(* IEC 61131-3 sources: STAR-PLC-Agent/results/raw/six_task_fullflow_20261114/PUB016/generation/sim_00, 1 file *)

(* ---- test_program.st ---- *)
PROGRAM PLC_PRG
VAR
 BenchStep : UDINT := 0;
 BenchCalls : UDINT := 0;
 BenchDone : BOOL := FALSE;
 BenchUut0 : FB_Task;
 BenchUut1 : FB_Task;
 TraceIn_processLength : ARRAY[0..12] OF USINT;
 TraceIn_sensor1 : ARRAY[0..12] OF BOOL;
 TraceIn_sensor2 : ARRAY[0..12] OF BOOL;
 TraceIn_sensor3 : ARRAY[0..12] OF BOOL;
 TraceIn_sensor4 : ARRAY[0..12] OF BOOL;
 TraceIn_sensor5 : ARRAY[0..12] OF BOOL;
 TraceIn_station1Start : ARRAY[0..12] OF BOOL;
 TraceIn_station2Complete : ARRAY[0..12] OF BOOL;
 TraceIn_station3Complete : ARRAY[0..12] OF BOOL;
 TraceIn_station4Complete : ARRAY[0..12] OF BOOL;
 TraceIn_processSequence_1 : ARRAY[0..12] OF USINT;
 TraceIn_processSequence_2 : ARRAY[0..12] OF USINT;
 TraceIn_processSequence_3 : ARRAY[0..12] OF USINT;
 TraceIn_processSequence_4 : ARRAY[0..12] OF USINT;
 TraceIn_processSequence_5 : ARRAY[0..12] OF USINT;
 TraceIn_processSequence_6 : ARRAY[0..12] OF USINT;
 TraceIn_processSequence_7 : ARRAY[0..12] OF USINT;
 TraceIn_processSequence_8 : ARRAY[0..12] OF USINT;
 TraceOut_conveyorLeft : ARRAY[0..12] OF BOOL;
 TraceOut_conveyorRight : ARRAY[0..12] OF BOOL;
END_VAR

IF NOT BenchDone THEN
 CASE BenchStep OF
 0:
   BenchUut0.processLength := USINT#2;
   BenchUut0.sensor1 := TRUE;
   BenchUut0.sensor2 := FALSE;
   BenchUut0.sensor3 := FALSE;
   BenchUut0.sensor4 := FALSE;
   BenchUut0.sensor5 := FALSE;
   BenchUut0.station1Start := FALSE;
   BenchUut0.station2Complete := FALSE;
   BenchUut0.station3Complete := FALSE;
   BenchUut0.station4Complete := FALSE;
   BenchUut0.processSequence[1] := USINT#2;
   BenchUut0.processSequence[2] := USINT#5;
   BenchUut0.processSequence[3] := USINT#0;
   BenchUut0.processSequence[4] := USINT#0;
   BenchUut0.processSequence[5] := USINT#0;
   BenchUut0.processSequence[6] := USINT#0;
   BenchUut0.processSequence[7] := USINT#0;
   BenchUut0.processSequence[8] := USINT#0;
   TraceIn_processLength[0] := BenchUut0.processLength;
   TraceIn_sensor1[0] := BenchUut0.sensor1;
   TraceIn_sensor2[0] := BenchUut0.sensor2;
   TraceIn_sensor3[0] := BenchUut0.sensor3;
   TraceIn_sensor4[0] := BenchUut0.sensor4;
   TraceIn_sensor5[0] := BenchUut0.sensor5;
   TraceIn_station1Start[0] := BenchUut0.station1Start;
   TraceIn_station2Complete[0] := BenchUut0.station2Complete;
   TraceIn_station3Complete[0] := BenchUut0.station3Complete;
   TraceIn_station4Complete[0] := BenchUut0.station4Complete;
   TraceIn_processSequence_1[0] := BenchUut0.processSequence[1];
   TraceIn_processSequence_2[0] := BenchUut0.processSequence[2];
   TraceIn_processSequence_3[0] := BenchUut0.processSequence[3];
   TraceIn_processSequence_4[0] := BenchUut0.processSequence[4];
   TraceIn_processSequence_5[0] := BenchUut0.processSequence[5];
   TraceIn_processSequence_6[0] := BenchUut0.processSequence[6];
   TraceIn_processSequence_7[0] := BenchUut0.processSequence[7];
   TraceIn_processSequence_8[0] := BenchUut0.processSequence[8];
   BenchUut0();
   TraceOut_conveyorLeft[0] := BenchUut0.conveyorLeft;
   TraceOut_conveyorRight[0] := BenchUut0.conveyorRight;
   BenchCalls := BenchCalls + 1;
 1:
   BenchUut0.processLength := USINT#2;
   BenchUut0.sensor1 := TRUE;
   BenchUut0.sensor2 := FALSE;
   BenchUut0.sensor3 := FALSE;
   BenchUut0.sensor4 := FALSE;
   BenchUut0.sensor5 := FALSE;
   BenchUut0.station1Start := TRUE;
   BenchUut0.station2Complete := FALSE;
   BenchUut0.station3Complete := FALSE;
   BenchUut0.station4Complete := FALSE;
   BenchUut0.processSequence[1] := USINT#2;
   BenchUut0.processSequence[2] := USINT#5;
   BenchUut0.processSequence[3] := USINT#0;
   BenchUut0.processSequence[4] := USINT#0;
   BenchUut0.processSequence[5] := USINT#0;
   BenchUut0.processSequence[6] := USINT#0;
   BenchUut0.processSequence[7] := USINT#0;
   BenchUut0.processSequence[8] := USINT#0;
   TraceIn_processLength[1] := BenchUut0.processLength;
   TraceIn_sensor1[1] := BenchUut0.sensor1;
   TraceIn_sensor2[1] := BenchUut0.sensor2;
   TraceIn_sensor3[1] := BenchUut0.sensor3;
   TraceIn_sensor4[1] := BenchUut0.sensor4;
   TraceIn_sensor5[1] := BenchUut0.sensor5;
   TraceIn_station1Start[1] := BenchUut0.station1Start;
   TraceIn_station2Complete[1] := BenchUut0.station2Complete;
   TraceIn_station3Complete[1] := BenchUut0.station3Complete;
   TraceIn_station4Complete[1] := BenchUut0.station4Complete;
   TraceIn_processSequence_1[1] := BenchUut0.processSequence[1];
   TraceIn_processSequence_2[1] := BenchUut0.processSequence[2];
   TraceIn_processSequence_3[1] := BenchUut0.processSequence[3];
   TraceIn_processSequence_4[1] := BenchUut0.processSequence[4];
   TraceIn_processSequence_5[1] := BenchUut0.processSequence[5];
   TraceIn_processSequence_6[1] := BenchUut0.processSequence[6];
   TraceIn_processSequence_7[1] := BenchUut0.processSequence[7];
   TraceIn_processSequence_8[1] := BenchUut0.processSequence[8];
   BenchUut0();
   TraceOut_conveyorLeft[1] := BenchUut0.conveyorLeft;
   TraceOut_conveyorRight[1] := BenchUut0.conveyorRight;
   BenchCalls := BenchCalls + 1;
 2:
   BenchUut0.processLength := USINT#2;
   BenchUut0.sensor1 := TRUE;
   BenchUut0.sensor2 := TRUE;
   BenchUut0.sensor3 := FALSE;
   BenchUut0.sensor4 := FALSE;
   BenchUut0.sensor5 := FALSE;
   BenchUut0.station1Start := FALSE;
   BenchUut0.station2Complete := FALSE;
   BenchUut0.station3Complete := FALSE;
   BenchUut0.station4Complete := FALSE;
   BenchUut0.processSequence[1] := USINT#2;
   BenchUut0.processSequence[2] := USINT#5;
   BenchUut0.processSequence[3] := USINT#0;
   BenchUut0.processSequence[4] := USINT#0;
   BenchUut0.processSequence[5] := USINT#0;
   BenchUut0.processSequence[6] := USINT#0;
   BenchUut0.processSequence[7] := USINT#0;
   BenchUut0.processSequence[8] := USINT#0;
   TraceIn_processLength[2] := BenchUut0.processLength;
   TraceIn_sensor1[2] := BenchUut0.sensor1;
   TraceIn_sensor2[2] := BenchUut0.sensor2;
   TraceIn_sensor3[2] := BenchUut0.sensor3;
   TraceIn_sensor4[2] := BenchUut0.sensor4;
   TraceIn_sensor5[2] := BenchUut0.sensor5;
   TraceIn_station1Start[2] := BenchUut0.station1Start;
   TraceIn_station2Complete[2] := BenchUut0.station2Complete;
   TraceIn_station3Complete[2] := BenchUut0.station3Complete;
   TraceIn_station4Complete[2] := BenchUut0.station4Complete;
   TraceIn_processSequence_1[2] := BenchUut0.processSequence[1];
   TraceIn_processSequence_2[2] := BenchUut0.processSequence[2];
   TraceIn_processSequence_3[2] := BenchUut0.processSequence[3];
   TraceIn_processSequence_4[2] := BenchUut0.processSequence[4];
   TraceIn_processSequence_5[2] := BenchUut0.processSequence[5];
   TraceIn_processSequence_6[2] := BenchUut0.processSequence[6];
   TraceIn_processSequence_7[2] := BenchUut0.processSequence[7];
   TraceIn_processSequence_8[2] := BenchUut0.processSequence[8];
   BenchUut0();
   TraceOut_conveyorLeft[2] := BenchUut0.conveyorLeft;
   TraceOut_conveyorRight[2] := BenchUut0.conveyorRight;
   BenchCalls := BenchCalls + 1;
 3:
   BenchUut0.processLength := USINT#2;
   BenchUut0.sensor1 := TRUE;
   BenchUut0.sensor2 := TRUE;
   BenchUut0.sensor3 := FALSE;
   BenchUut0.sensor4 := FALSE;
   BenchUut0.sensor5 := FALSE;
   BenchUut0.station1Start := FALSE;
   BenchUut0.station2Complete := TRUE;
   BenchUut0.station3Complete := FALSE;
   BenchUut0.station4Complete := FALSE;
   BenchUut0.processSequence[1] := USINT#2;
   BenchUut0.processSequence[2] := USINT#5;
   BenchUut0.processSequence[3] := USINT#0;
   BenchUut0.processSequence[4] := USINT#0;
   BenchUut0.processSequence[5] := USINT#0;
   BenchUut0.processSequence[6] := USINT#0;
   BenchUut0.processSequence[7] := USINT#0;
   BenchUut0.processSequence[8] := USINT#0;
   TraceIn_processLength[3] := BenchUut0.processLength;
   TraceIn_sensor1[3] := BenchUut0.sensor1;
   TraceIn_sensor2[3] := BenchUut0.sensor2;
   TraceIn_sensor3[3] := BenchUut0.sensor3;
   TraceIn_sensor4[3] := BenchUut0.sensor4;
   TraceIn_sensor5[3] := BenchUut0.sensor5;
   TraceIn_station1Start[3] := BenchUut0.station1Start;
   TraceIn_station2Complete[3] := BenchUut0.station2Complete;
   TraceIn_station3Complete[3] := BenchUut0.station3Complete;
   TraceIn_station4Complete[3] := BenchUut0.station4Complete;
   TraceIn_processSequence_1[3] := BenchUut0.processSequence[1];
   TraceIn_processSequence_2[3] := BenchUut0.processSequence[2];
   TraceIn_processSequence_3[3] := BenchUut0.processSequence[3];
   TraceIn_processSequence_4[3] := BenchUut0.processSequence[4];
   TraceIn_processSequence_5[3] := BenchUut0.processSequence[5];
   TraceIn_processSequence_6[3] := BenchUut0.processSequence[6];
   TraceIn_processSequence_7[3] := BenchUut0.processSequence[7];
   TraceIn_processSequence_8[3] := BenchUut0.processSequence[8];
   BenchUut0();
   TraceOut_conveyorLeft[3] := BenchUut0.conveyorLeft;
   TraceOut_conveyorRight[3] := BenchUut0.conveyorRight;
   BenchCalls := BenchCalls + 1;
 4:
   BenchUut0.processLength := USINT#2;
   BenchUut0.sensor1 := FALSE;
   BenchUut0.sensor2 := FALSE;
   BenchUut0.sensor3 := FALSE;
   BenchUut0.sensor4 := FALSE;
   BenchUut0.sensor5 := FALSE;
   BenchUut0.station1Start := FALSE;
   BenchUut0.station2Complete := FALSE;
   BenchUut0.station3Complete := FALSE;
   BenchUut0.station4Complete := FALSE;
   BenchUut0.processSequence[1] := USINT#2;
   BenchUut0.processSequence[2] := USINT#5;
   BenchUut0.processSequence[3] := USINT#0;
   BenchUut0.processSequence[4] := USINT#0;
   BenchUut0.processSequence[5] := USINT#0;
   BenchUut0.processSequence[6] := USINT#0;
   BenchUut0.processSequence[7] := USINT#0;
   BenchUut0.processSequence[8] := USINT#0;
   TraceIn_processLength[4] := BenchUut0.processLength;
   TraceIn_sensor1[4] := BenchUut0.sensor1;
   TraceIn_sensor2[4] := BenchUut0.sensor2;
   TraceIn_sensor3[4] := BenchUut0.sensor3;
   TraceIn_sensor4[4] := BenchUut0.sensor4;
   TraceIn_sensor5[4] := BenchUut0.sensor5;
   TraceIn_station1Start[4] := BenchUut0.station1Start;
   TraceIn_station2Complete[4] := BenchUut0.station2Complete;
   TraceIn_station3Complete[4] := BenchUut0.station3Complete;
   TraceIn_station4Complete[4] := BenchUut0.station4Complete;
   TraceIn_processSequence_1[4] := BenchUut0.processSequence[1];
   TraceIn_processSequence_2[4] := BenchUut0.processSequence[2];
   TraceIn_processSequence_3[4] := BenchUut0.processSequence[3];
   TraceIn_processSequence_4[4] := BenchUut0.processSequence[4];
   TraceIn_processSequence_5[4] := BenchUut0.processSequence[5];
   TraceIn_processSequence_6[4] := BenchUut0.processSequence[6];
   TraceIn_processSequence_7[4] := BenchUut0.processSequence[7];
   TraceIn_processSequence_8[4] := BenchUut0.processSequence[8];
   BenchUut0();
   TraceOut_conveyorLeft[4] := BenchUut0.conveyorLeft;
   TraceOut_conveyorRight[4] := BenchUut0.conveyorRight;
   BenchCalls := BenchCalls + 1;
 5:
   BenchUut0.processLength := USINT#2;
   BenchUut0.sensor1 := FALSE;
   BenchUut0.sensor2 := FALSE;
   BenchUut0.sensor3 := FALSE;
   BenchUut0.sensor4 := FALSE;
   BenchUut0.sensor5 := TRUE;
   BenchUut0.station1Start := FALSE;
   BenchUut0.station2Complete := FALSE;
   BenchUut0.station3Complete := FALSE;
   BenchUut0.station4Complete := FALSE;
   BenchUut0.processSequence[1] := USINT#2;
   BenchUut0.processSequence[2] := USINT#5;
   BenchUut0.processSequence[3] := USINT#0;
   BenchUut0.processSequence[4] := USINT#0;
   BenchUut0.processSequence[5] := USINT#0;
   BenchUut0.processSequence[6] := USINT#0;
   BenchUut0.processSequence[7] := USINT#0;
   BenchUut0.processSequence[8] := USINT#0;
   TraceIn_processLength[5] := BenchUut0.processLength;
   TraceIn_sensor1[5] := BenchUut0.sensor1;
   TraceIn_sensor2[5] := BenchUut0.sensor2;
   TraceIn_sensor3[5] := BenchUut0.sensor3;
   TraceIn_sensor4[5] := BenchUut0.sensor4;
   TraceIn_sensor5[5] := BenchUut0.sensor5;
   TraceIn_station1Start[5] := BenchUut0.station1Start;
   TraceIn_station2Complete[5] := BenchUut0.station2Complete;
   TraceIn_station3Complete[5] := BenchUut0.station3Complete;
   TraceIn_station4Complete[5] := BenchUut0.station4Complete;
   TraceIn_processSequence_1[5] := BenchUut0.processSequence[1];
   TraceIn_processSequence_2[5] := BenchUut0.processSequence[2];
   TraceIn_processSequence_3[5] := BenchUut0.processSequence[3];
   TraceIn_processSequence_4[5] := BenchUut0.processSequence[4];
   TraceIn_processSequence_5[5] := BenchUut0.processSequence[5];
   TraceIn_processSequence_6[5] := BenchUut0.processSequence[6];
   TraceIn_processSequence_7[5] := BenchUut0.processSequence[7];
   TraceIn_processSequence_8[5] := BenchUut0.processSequence[8];
   BenchUut0();
   TraceOut_conveyorLeft[5] := BenchUut0.conveyorLeft;
   TraceOut_conveyorRight[5] := BenchUut0.conveyorRight;
   BenchCalls := BenchCalls + 1;
 6:
   BenchUut1.processLength := USINT#3;
   BenchUut1.sensor1 := TRUE;
   BenchUut1.sensor2 := FALSE;
   BenchUut1.sensor3 := FALSE;
   BenchUut1.sensor4 := FALSE;
   BenchUut1.sensor5 := FALSE;
   BenchUut1.station1Start := FALSE;
   BenchUut1.station2Complete := FALSE;
   BenchUut1.station3Complete := FALSE;
   BenchUut1.station4Complete := FALSE;
   BenchUut1.processSequence[1] := USINT#2;
   BenchUut1.processSequence[2] := USINT#2;
   BenchUut1.processSequence[3] := USINT#5;
   BenchUut1.processSequence[4] := USINT#0;
   BenchUut1.processSequence[5] := USINT#0;
   BenchUut1.processSequence[6] := USINT#0;
   BenchUut1.processSequence[7] := USINT#0;
   BenchUut1.processSequence[8] := USINT#0;
   TraceIn_processLength[6] := BenchUut1.processLength;
   TraceIn_sensor1[6] := BenchUut1.sensor1;
   TraceIn_sensor2[6] := BenchUut1.sensor2;
   TraceIn_sensor3[6] := BenchUut1.sensor3;
   TraceIn_sensor4[6] := BenchUut1.sensor4;
   TraceIn_sensor5[6] := BenchUut1.sensor5;
   TraceIn_station1Start[6] := BenchUut1.station1Start;
   TraceIn_station2Complete[6] := BenchUut1.station2Complete;
   TraceIn_station3Complete[6] := BenchUut1.station3Complete;
   TraceIn_station4Complete[6] := BenchUut1.station4Complete;
   TraceIn_processSequence_1[6] := BenchUut1.processSequence[1];
   TraceIn_processSequence_2[6] := BenchUut1.processSequence[2];
   TraceIn_processSequence_3[6] := BenchUut1.processSequence[3];
   TraceIn_processSequence_4[6] := BenchUut1.processSequence[4];
   TraceIn_processSequence_5[6] := BenchUut1.processSequence[5];
   TraceIn_processSequence_6[6] := BenchUut1.processSequence[6];
   TraceIn_processSequence_7[6] := BenchUut1.processSequence[7];
   TraceIn_processSequence_8[6] := BenchUut1.processSequence[8];
   BenchUut1();
   TraceOut_conveyorLeft[6] := BenchUut1.conveyorLeft;
   TraceOut_conveyorRight[6] := BenchUut1.conveyorRight;
   BenchCalls := BenchCalls + 1;
 7:
   BenchUut1.processLength := USINT#3;
   BenchUut1.sensor1 := TRUE;
   BenchUut1.sensor2 := FALSE;
   BenchUut1.sensor3 := FALSE;
   BenchUut1.sensor4 := FALSE;
   BenchUut1.sensor5 := FALSE;
   BenchUut1.station1Start := TRUE;
   BenchUut1.station2Complete := FALSE;
   BenchUut1.station3Complete := FALSE;
   BenchUut1.station4Complete := FALSE;
   BenchUut1.processSequence[1] := USINT#2;
   BenchUut1.processSequence[2] := USINT#2;
   BenchUut1.processSequence[3] := USINT#5;
   BenchUut1.processSequence[4] := USINT#0;
   BenchUut1.processSequence[5] := USINT#0;
   BenchUut1.processSequence[6] := USINT#0;
   BenchUut1.processSequence[7] := USINT#0;
   BenchUut1.processSequence[8] := USINT#0;
   TraceIn_processLength[7] := BenchUut1.processLength;
   TraceIn_sensor1[7] := BenchUut1.sensor1;
   TraceIn_sensor2[7] := BenchUut1.sensor2;
   TraceIn_sensor3[7] := BenchUut1.sensor3;
   TraceIn_sensor4[7] := BenchUut1.sensor4;
   TraceIn_sensor5[7] := BenchUut1.sensor5;
   TraceIn_station1Start[7] := BenchUut1.station1Start;
   TraceIn_station2Complete[7] := BenchUut1.station2Complete;
   TraceIn_station3Complete[7] := BenchUut1.station3Complete;
   TraceIn_station4Complete[7] := BenchUut1.station4Complete;
   TraceIn_processSequence_1[7] := BenchUut1.processSequence[1];
   TraceIn_processSequence_2[7] := BenchUut1.processSequence[2];
   TraceIn_processSequence_3[7] := BenchUut1.processSequence[3];
   TraceIn_processSequence_4[7] := BenchUut1.processSequence[4];
   TraceIn_processSequence_5[7] := BenchUut1.processSequence[5];
   TraceIn_processSequence_6[7] := BenchUut1.processSequence[6];
   TraceIn_processSequence_7[7] := BenchUut1.processSequence[7];
   TraceIn_processSequence_8[7] := BenchUut1.processSequence[8];
   BenchUut1();
   TraceOut_conveyorLeft[7] := BenchUut1.conveyorLeft;
   TraceOut_conveyorRight[7] := BenchUut1.conveyorRight;
   BenchCalls := BenchCalls + 1;
 8:
   BenchUut1.processLength := USINT#3;
   BenchUut1.sensor1 := TRUE;
   BenchUut1.sensor2 := TRUE;
   BenchUut1.sensor3 := FALSE;
   BenchUut1.sensor4 := FALSE;
   BenchUut1.sensor5 := FALSE;
   BenchUut1.station1Start := FALSE;
   BenchUut1.station2Complete := FALSE;
   BenchUut1.station3Complete := FALSE;
   BenchUut1.station4Complete := FALSE;
   BenchUut1.processSequence[1] := USINT#2;
   BenchUut1.processSequence[2] := USINT#2;
   BenchUut1.processSequence[3] := USINT#5;
   BenchUut1.processSequence[4] := USINT#0;
   BenchUut1.processSequence[5] := USINT#0;
   BenchUut1.processSequence[6] := USINT#0;
   BenchUut1.processSequence[7] := USINT#0;
   BenchUut1.processSequence[8] := USINT#0;
   TraceIn_processLength[8] := BenchUut1.processLength;
   TraceIn_sensor1[8] := BenchUut1.sensor1;
   TraceIn_sensor2[8] := BenchUut1.sensor2;
   TraceIn_sensor3[8] := BenchUut1.sensor3;
   TraceIn_sensor4[8] := BenchUut1.sensor4;
   TraceIn_sensor5[8] := BenchUut1.sensor5;
   TraceIn_station1Start[8] := BenchUut1.station1Start;
   TraceIn_station2Complete[8] := BenchUut1.station2Complete;
   TraceIn_station3Complete[8] := BenchUut1.station3Complete;
   TraceIn_station4Complete[8] := BenchUut1.station4Complete;
   TraceIn_processSequence_1[8] := BenchUut1.processSequence[1];
   TraceIn_processSequence_2[8] := BenchUut1.processSequence[2];
   TraceIn_processSequence_3[8] := BenchUut1.processSequence[3];
   TraceIn_processSequence_4[8] := BenchUut1.processSequence[4];
   TraceIn_processSequence_5[8] := BenchUut1.processSequence[5];
   TraceIn_processSequence_6[8] := BenchUut1.processSequence[6];
   TraceIn_processSequence_7[8] := BenchUut1.processSequence[7];
   TraceIn_processSequence_8[8] := BenchUut1.processSequence[8];
   BenchUut1();
   TraceOut_conveyorLeft[8] := BenchUut1.conveyorLeft;
   TraceOut_conveyorRight[8] := BenchUut1.conveyorRight;
   BenchCalls := BenchCalls + 1;
 9:
   BenchUut1.processLength := USINT#3;
   BenchUut1.sensor1 := TRUE;
   BenchUut1.sensor2 := TRUE;
   BenchUut1.sensor3 := FALSE;
   BenchUut1.sensor4 := FALSE;
   BenchUut1.sensor5 := FALSE;
   BenchUut1.station1Start := FALSE;
   BenchUut1.station2Complete := TRUE;
   BenchUut1.station3Complete := FALSE;
   BenchUut1.station4Complete := FALSE;
   BenchUut1.processSequence[1] := USINT#2;
   BenchUut1.processSequence[2] := USINT#2;
   BenchUut1.processSequence[3] := USINT#5;
   BenchUut1.processSequence[4] := USINT#0;
   BenchUut1.processSequence[5] := USINT#0;
   BenchUut1.processSequence[6] := USINT#0;
   BenchUut1.processSequence[7] := USINT#0;
   BenchUut1.processSequence[8] := USINT#0;
   TraceIn_processLength[9] := BenchUut1.processLength;
   TraceIn_sensor1[9] := BenchUut1.sensor1;
   TraceIn_sensor2[9] := BenchUut1.sensor2;
   TraceIn_sensor3[9] := BenchUut1.sensor3;
   TraceIn_sensor4[9] := BenchUut1.sensor4;
   TraceIn_sensor5[9] := BenchUut1.sensor5;
   TraceIn_station1Start[9] := BenchUut1.station1Start;
   TraceIn_station2Complete[9] := BenchUut1.station2Complete;
   TraceIn_station3Complete[9] := BenchUut1.station3Complete;
   TraceIn_station4Complete[9] := BenchUut1.station4Complete;
   TraceIn_processSequence_1[9] := BenchUut1.processSequence[1];
   TraceIn_processSequence_2[9] := BenchUut1.processSequence[2];
   TraceIn_processSequence_3[9] := BenchUut1.processSequence[3];
   TraceIn_processSequence_4[9] := BenchUut1.processSequence[4];
   TraceIn_processSequence_5[9] := BenchUut1.processSequence[5];
   TraceIn_processSequence_6[9] := BenchUut1.processSequence[6];
   TraceIn_processSequence_7[9] := BenchUut1.processSequence[7];
   TraceIn_processSequence_8[9] := BenchUut1.processSequence[8];
   BenchUut1();
   TraceOut_conveyorLeft[9] := BenchUut1.conveyorLeft;
   TraceOut_conveyorRight[9] := BenchUut1.conveyorRight;
   BenchCalls := BenchCalls + 1;
 10:
   BenchUut1.processLength := USINT#3;
   BenchUut1.sensor1 := TRUE;
   BenchUut1.sensor2 := TRUE;
   BenchUut1.sensor3 := FALSE;
   BenchUut1.sensor4 := FALSE;
   BenchUut1.sensor5 := FALSE;
   BenchUut1.station1Start := FALSE;
   BenchUut1.station2Complete := FALSE;
   BenchUut1.station3Complete := FALSE;
   BenchUut1.station4Complete := FALSE;
   BenchUut1.processSequence[1] := USINT#2;
   BenchUut1.processSequence[2] := USINT#2;
   BenchUut1.processSequence[3] := USINT#5;
   BenchUut1.processSequence[4] := USINT#0;
   BenchUut1.processSequence[5] := USINT#0;
   BenchUut1.processSequence[6] := USINT#0;
   BenchUut1.processSequence[7] := USINT#0;
   BenchUut1.processSequence[8] := USINT#0;
   TraceIn_processLength[10] := BenchUut1.processLength;
   TraceIn_sensor1[10] := BenchUut1.sensor1;
   TraceIn_sensor2[10] := BenchUut1.sensor2;
   TraceIn_sensor3[10] := BenchUut1.sensor3;
   TraceIn_sensor4[10] := BenchUut1.sensor4;
   TraceIn_sensor5[10] := BenchUut1.sensor5;
   TraceIn_station1Start[10] := BenchUut1.station1Start;
   TraceIn_station2Complete[10] := BenchUut1.station2Complete;
   TraceIn_station3Complete[10] := BenchUut1.station3Complete;
   TraceIn_station4Complete[10] := BenchUut1.station4Complete;
   TraceIn_processSequence_1[10] := BenchUut1.processSequence[1];
   TraceIn_processSequence_2[10] := BenchUut1.processSequence[2];
   TraceIn_processSequence_3[10] := BenchUut1.processSequence[3];
   TraceIn_processSequence_4[10] := BenchUut1.processSequence[4];
   TraceIn_processSequence_5[10] := BenchUut1.processSequence[5];
   TraceIn_processSequence_6[10] := BenchUut1.processSequence[6];
   TraceIn_processSequence_7[10] := BenchUut1.processSequence[7];
   TraceIn_processSequence_8[10] := BenchUut1.processSequence[8];
   BenchUut1();
   TraceOut_conveyorLeft[10] := BenchUut1.conveyorLeft;
   TraceOut_conveyorRight[10] := BenchUut1.conveyorRight;
   BenchCalls := BenchCalls + 1;
 11:
   BenchUut1.processLength := USINT#3;
   BenchUut1.sensor1 := TRUE;
   BenchUut1.sensor2 := TRUE;
   BenchUut1.sensor3 := FALSE;
   BenchUut1.sensor4 := FALSE;
   BenchUut1.sensor5 := FALSE;
   BenchUut1.station1Start := FALSE;
   BenchUut1.station2Complete := TRUE;
   BenchUut1.station3Complete := FALSE;
   BenchUut1.station4Complete := FALSE;
   BenchUut1.processSequence[1] := USINT#2;
   BenchUut1.processSequence[2] := USINT#2;
   BenchUut1.processSequence[3] := USINT#5;
   BenchUut1.processSequence[4] := USINT#0;
   BenchUut1.processSequence[5] := USINT#0;
   BenchUut1.processSequence[6] := USINT#0;
   BenchUut1.processSequence[7] := USINT#0;
   BenchUut1.processSequence[8] := USINT#0;
   TraceIn_processLength[11] := BenchUut1.processLength;
   TraceIn_sensor1[11] := BenchUut1.sensor1;
   TraceIn_sensor2[11] := BenchUut1.sensor2;
   TraceIn_sensor3[11] := BenchUut1.sensor3;
   TraceIn_sensor4[11] := BenchUut1.sensor4;
   TraceIn_sensor5[11] := BenchUut1.sensor5;
   TraceIn_station1Start[11] := BenchUut1.station1Start;
   TraceIn_station2Complete[11] := BenchUut1.station2Complete;
   TraceIn_station3Complete[11] := BenchUut1.station3Complete;
   TraceIn_station4Complete[11] := BenchUut1.station4Complete;
   TraceIn_processSequence_1[11] := BenchUut1.processSequence[1];
   TraceIn_processSequence_2[11] := BenchUut1.processSequence[2];
   TraceIn_processSequence_3[11] := BenchUut1.processSequence[3];
   TraceIn_processSequence_4[11] := BenchUut1.processSequence[4];
   TraceIn_processSequence_5[11] := BenchUut1.processSequence[5];
   TraceIn_processSequence_6[11] := BenchUut1.processSequence[6];
   TraceIn_processSequence_7[11] := BenchUut1.processSequence[7];
   TraceIn_processSequence_8[11] := BenchUut1.processSequence[8];
   BenchUut1();
   TraceOut_conveyorLeft[11] := BenchUut1.conveyorLeft;
   TraceOut_conveyorRight[11] := BenchUut1.conveyorRight;
   BenchCalls := BenchCalls + 1;
 12:
   BenchUut1.processLength := USINT#3;
   BenchUut1.sensor1 := FALSE;
   BenchUut1.sensor2 := FALSE;
   BenchUut1.sensor3 := FALSE;
   BenchUut1.sensor4 := FALSE;
   BenchUut1.sensor5 := TRUE;
   BenchUut1.station1Start := FALSE;
   BenchUut1.station2Complete := FALSE;
   BenchUut1.station3Complete := FALSE;
   BenchUut1.station4Complete := FALSE;
   BenchUut1.processSequence[1] := USINT#2;
   BenchUut1.processSequence[2] := USINT#2;
   BenchUut1.processSequence[3] := USINT#5;
   BenchUut1.processSequence[4] := USINT#0;
   BenchUut1.processSequence[5] := USINT#0;
   BenchUut1.processSequence[6] := USINT#0;
   BenchUut1.processSequence[7] := USINT#0;
   BenchUut1.processSequence[8] := USINT#0;
   TraceIn_processLength[12] := BenchUut1.processLength;
   TraceIn_sensor1[12] := BenchUut1.sensor1;
   TraceIn_sensor2[12] := BenchUut1.sensor2;
   TraceIn_sensor3[12] := BenchUut1.sensor3;
   TraceIn_sensor4[12] := BenchUut1.sensor4;
   TraceIn_sensor5[12] := BenchUut1.sensor5;
   TraceIn_station1Start[12] := BenchUut1.station1Start;
   TraceIn_station2Complete[12] := BenchUut1.station2Complete;
   TraceIn_station3Complete[12] := BenchUut1.station3Complete;
   TraceIn_station4Complete[12] := BenchUut1.station4Complete;
   TraceIn_processSequence_1[12] := BenchUut1.processSequence[1];
   TraceIn_processSequence_2[12] := BenchUut1.processSequence[2];
   TraceIn_processSequence_3[12] := BenchUut1.processSequence[3];
   TraceIn_processSequence_4[12] := BenchUut1.processSequence[4];
   TraceIn_processSequence_5[12] := BenchUut1.processSequence[5];
   TraceIn_processSequence_6[12] := BenchUut1.processSequence[6];
   TraceIn_processSequence_7[12] := BenchUut1.processSequence[7];
   TraceIn_processSequence_8[12] := BenchUut1.processSequence[8];
   BenchUut1();
   TraceOut_conveyorLeft[12] := BenchUut1.conveyorLeft;
   TraceOut_conveyorRight[12] := BenchUut1.conveyorRight;
   BenchCalls := BenchCalls + 1;
 END_CASE;
 BenchStep := BenchStep + 1;
 IF BenchStep >= 13 THEN BenchDone := TRUE; END_IF;
END_IF;
END_PROGRAM
